// TwinCAT 3 PLC project Untitled1
// ProgramVersion: 3.1.4026.25
// libraries:
//   Tc2_Standard, * (Beckhoff Automation GmbH)
//   Tc2_System, * (Beckhoff Automation GmbH)
// project tree:
//   GVLs/ GVL.TcGVL
//   / PlcTask.TcTTO
//   POUs/ MAIN.TcPOU
// real-time tasks:
//   TASK PlcTask: cycle T#10ms, priority 20, ADS port 350
// motion (NC):
//   TASK NC-Task 1 SAF: cycle T#2ms, priority 4, ADS port 501
//   TASK NC-Task 1 SVB: cycle T#10ms, priority 8, ADS port 511
//   AXIS Axis 1 (id 1)
//     OtherSettings: AllowMotionCmdToSlave=true
//     encoder EncType=8
//       EncPara: MaxCount=#xffffffff
//     drive DrvType=9
//       DrvPara: MaxCount=#xffffffff, DriveControlDWord=#x00030000
//         Analog: VeloScale=6, TorqueSetpointScale=10, ScaleFactorActTorque=0.1
//         TimeComp: TaskDelayCycles=1
//     controller CtrType=1
//       CtrPara: PriorControlFactor=1
//         Observer: BandWidth=20
//   AXIS Axis 2 (id 2)
//     OtherSettings: AllowMotionCmdToSlave=true
//     encoder EncType=8
//       EncPara: MaxCount=#xffffffff
//     drive DrvType=9
//       DrvPara: MaxCount=#xffffffff, DriveControlDWord=#x00030000
//         Analog: VeloScale=6, TorqueSetpointScale=10, ScaleFactorActTorque=0.1
//         TimeComp: TaskDelayCycles=1
//     controller CtrType=1
//       CtrPara: PriorControlFactor=1
//         Observer: BandWidth=20
// I/O:
//   DEVICE Device 1 (EtherCAT), AmsNetId 192.168.0.5.2.1
//     Box 1 (CU1128) [CU1128 6x EtherCAT junction]
//       Box 10 (EP1018-0001) [EP1018-0001 8 Ch. Dig. Input 24V, 10µs, M8]
//       Box 11 (EP1018-0001) [EP1018-0001 8 Ch. Dig. Input 24V, 10µs, M8]
//       Box 12 (EP1018-0001) [EP1018-0001 8 Ch. Dig. Input 24V, 10µs, M8]
//       Box 13 (EP2028-0001) [EP2028-0001 8 Ch. Dig. Output 24V, 2A, M8]
//       Box 14 (EP2028-0001) [EP2028-0001 8 Ch. Dig. Output 24V, 2A, M8]
//       Term 7 (EK1100-0030) [EK1100-0030 EtherCAT Coupler (2A E-Bus, 4kV galv. iso.)]
//         Term 8 (EL1809) [EL1809 16Ch. Dig. Input 24V, 3ms]
//         Term 9 (EL2809) [EL2809 16Ch. Dig. Output 24V, 0.5A]
//       Term 4 (EK1100-0030) [EK1100-0030 EtherCAT Coupler (2A E-Bus, 4kV galv. iso.)]
//         Term 5 (EL1809) [EL1809 16Ch. Dig. Input 24V, 3ms]
//         Term 6 (EL2809) [EL2809 16Ch. Dig. Output 24V, 0.5A]
//         Drive 15 (AX5206-0000-0011) [AX5206-0000-0011 EtherCAT Drive (SoE, 2 Ch.)]
//       Box 2 (CU1128-B) [CU1128 6x EtherCAT junction - Dev A]
//       Box 3 (CU1128-C) [CU1128 6x EtherCAT junction - Dev B]
// variable links:
//   NC-Task 1 SAF/Axes/Axis 1 <-> Device 1 (EtherCAT)/Box 1 (CU1128)/Term 4 (EK1100-0030)/Drive 15 (AX5206-0000-0011)
//     Drive/Inputs/In/nDcOutputTime <-> InfoData/DcOutputShift
//     Drive/Inputs/In/nState1 <-> AT 1/Drive status word @bit 8
//     Drive/Inputs/In/nState2 <-> AT 1/Drive status word
//     Drive/Inputs/In/nState4 @bit 1 <-> WcState/InputToggle
//     Drive/Inputs/In/nState4 <-> WcState/WcState
//     Drive/Outputs/Out/nCtrl1 <-> MDT 1/Master control word @bit 8
//     Drive/Outputs/Out/nDataOut2 <-> MDT 1/Velocity command value
//     Enc/Inputs/In/nDataIn1 <-> AT 1/Position feedback 1 value
//     Enc/Inputs/In/nDcInputTime <-> InfoData/DcInputShift
//     Enc/Inputs/In/nState4 @bit 1 <-> WcState/InputToggle
//     Enc/Inputs/In/nState4 <-> WcState/WcState
//   NC-Task 1 SAF/Axes/Axis 2 <-> Device 1 (EtherCAT)/Box 1 (CU1128)/Term 4 (EK1100-0030)/Drive 15 (AX5206-0000-0011)
//     Drive/Inputs/In/nDcOutputTime <-> InfoData/DcOutputShift
//     Drive/Inputs/In/nState1 <-> AT 2/Drive status word @bit 8
//     Drive/Inputs/In/nState2 <-> AT 2/Drive status word
//     Drive/Inputs/In/nState4 @bit 1 <-> WcState/InputToggle
//     Drive/Inputs/In/nState4 <-> WcState/WcState
//     Drive/Outputs/Out/nCtrl1 <-> MDT 2/Master control word @bit 8
//     Drive/Outputs/Out/nDataOut2 <-> MDT 2/Velocity command value
//     Enc/Inputs/In/nDataIn1 <-> AT 2/Position feedback 1 value
//     Enc/Inputs/In/nDcInputTime <-> InfoData/DcInputShift
//     Enc/Inputs/In/nState4 @bit 1 <-> WcState/InputToggle
//     Enc/Inputs/In/nState4 <-> WcState/WcState
//   Untitled1/Untitled1 Instance <-> Device 1 (EtherCAT)/Box 1 (CU1128)/Box 10 (EP1018-0001)
//     PlcTask Inputs/GVL.bZylAuswerferAS <-> Channel 1/Input
//     PlcTask Inputs/GVL.bZylAuswerferGS <-> Channel 2/Input
//     PlcTask Inputs/GVL.bZylSpannerAS <-> Channel 3/Input
//     PlcTask Inputs/GVL.bZylSpannerGS <-> Channel 4/Input
//     PlcTask Inputs/GVL.bZylWeicheAS <-> Channel 5/Input
//     PlcTask Inputs/GVL.bZylWeicheGS <-> Channel 6/Input
//   Untitled1/Untitled1 Instance <-> Device 1 (EtherCAT)/Box 1 (CU1128)/Box 11 (EP1018-0001)
//     PlcTask Inputs/GVL.bZylAuslaufAS <-> Channel 3/Input
//     PlcTask Inputs/GVL.bZylAuslaufGS <-> Channel 4/Input
//     PlcTask Inputs/GVL.bZylEinlaufAS <-> Channel 1/Input
//     PlcTask Inputs/GVL.bZylEinlaufGS <-> Channel 2/Input
//   Untitled1/Untitled1 Instance <-> Device 1 (EtherCAT)/Box 1 (CU1128)/Box 12 (EP1018-0001)
//     PlcTask Inputs/GVL.bLS_Auslauf <-> Channel 5/Input
//     PlcTask Inputs/GVL.bLS_Einlauf <-> Channel 1/Input
//     PlcTask Inputs/GVL.bServoAuslaufAS <-> Channel 7/Input
//     PlcTask Inputs/GVL.bServoAuslaufGS <-> Channel 8/Input
//     PlcTask Inputs/GVL.bServoAuslaufRast <-> Channel 6/Input
//     PlcTask Inputs/GVL.bServoEinlaufAS <-> Channel 3/Input
//     PlcTask Inputs/GVL.bServoEinlaufGS <-> Channel 4/Input
//     PlcTask Inputs/GVL.bServoEinlaufRast <-> Channel 2/Input
//   Untitled1/Untitled1 Instance <-> Device 1 (EtherCAT)/Box 1 (CU1128)/Box 13 (EP2028-0001)
//     PlcTask Outputs/GVL.bVentilAuswerferAS <-> Channel 1/Output
//     PlcTask Outputs/GVL.bVentilAuswerferGS <-> Channel 2/Output
//     PlcTask Outputs/GVL.bVentilSpannerAS <-> Channel 3/Output
//     PlcTask Outputs/GVL.bVentilSpannerGS <-> Channel 4/Output
//     PlcTask Outputs/GVL.bVentilWeicheAS <-> Channel 5/Output
//     PlcTask Outputs/GVL.bVentilWeicheGS <-> Channel 6/Output
//   Untitled1/Untitled1 Instance <-> Device 1 (EtherCAT)/Box 1 (CU1128)/Box 14 (EP2028-0001)
//     PlcTask Outputs/GVL.bVentilAusblasenAS <-> Channel 5/Output
//     PlcTask Outputs/GVL.bVentilAusblasenGS <-> Channel 6/Output
//     PlcTask Outputs/GVL.bVentilAuslaufAS <-> Channel 3/Output
//     PlcTask Outputs/GVL.bVentilAuslaufGS <-> Channel 4/Output
//     PlcTask Outputs/GVL.bVentilAuswurfBypAS <-> Channel 7/Output
//     PlcTask Outputs/GVL.bVentilAuswurfBypGS <-> Channel 8/Output
//     PlcTask Outputs/GVL.bVentilEinlaufAS <-> Channel 1/Output
//     PlcTask Outputs/GVL.bVentilEinlaufGS <-> Channel 2/Output
//   Untitled1/Untitled1 Instance <-> Device 1 (EtherCAT)/Box 1 (CU1128)/Term 4 (EK1100-0030)/Term 5 (EL1809)
//     PlcTask Inputs/GVL.bDruckschalter <-> Channel 1/Input
//     PlcTask Inputs/GVL.bNotHalt <-> Channel 2/Input
//   Untitled1/Untitled1 Instance <-> Device 1 (EtherCAT)/Box 1 (CU1128)/Term 4 (EK1100-0030)/Term 6 (EL2809)
//     PlcTask Outputs/GVL.bEntlueften <-> Channel 1/Output
//     PlcTask Outputs/GVL.bLaserEnable <-> Channel 2/Output
//   Untitled1/Untitled1 Instance <-> Device 1 (EtherCAT)/Box 1 (CU1128)/Term 7 (EK1100-0030)/Term 8 (EL1809)
//     PlcTask Inputs/GVL.bCW_Adb_coded <-> Channel 2/Input
//     PlcTask Inputs/GVL.bCW_Eready <-> Channel 1/Input
//     PlcTask Inputs/GVL.bCW_MarkInProgress <-> Channel 3/Input
//   Untitled1/Untitled1 Instance <-> Device 1 (EtherCAT)/Box 1 (CU1128)/Term 7 (EK1100-0030)/Term 9 (EL2809)
//     PlcTask Outputs/GVL.bCW_ERR_RESET <-> Channel 2/Output
//     PlcTask Outputs/GVL.bCW_Ex_GO <-> Channel 1/Output
//     PlcTask Outputs/GVL.bCW_STAT_REQ <-> Channel 4/Output
//     PlcTask Outputs/GVL.bCW_STOP <-> Channel 3/Output

CONFIGURATION Untitled1
    RESOURCE PLC ON TwinCAT3
        TASK PlcTask(INTERVAL := T#10ms, PRIORITY := 20);
        PROGRAM MAIN WITH PlcTask : MAIN;
    END_RESOURCE
END_CONFIGURATION

// ---- GVLs/GVL.TcGVL
{attribute 'qualified_only'}
VAR_GLOBAL
    // ==========================================
    // MAIN CONTROL CABINET (Schaltschrank)
    // ==========================================
    
    // Inputs (EL1809 - +MP-6K10)
    bDruckschalter         AT %I* : BOOL; // E0.0 Wartungseinheit Druckschalter[cite: 15, 25]
    bNotHalt               AT %I* : BOOL; // E0.1 Not-Halt betätigt[cite: 15, 18]
    
    // Outputs (EL2809 - +MP-6K20)
    bEntlueften            AT %Q* : BOOL; // A0.0 Wartungseinheit Entlüften[cite: 15, 25]
    bLaserEnable           AT %Q* : BOOL; // A0.1 LaserEnable[cite: 15, 18]

    // ==========================================
    // CW CONTROLLER
    // ==========================================
    
    // Inputs (EL1809 - +LS-7K10)
    bCW_Eready             AT %I* : BOOL; // E50.0 CW Eready[cite: 17]
    bCW_Adb_coded          AT %I* : BOOL; // E50.1 CW Adb coded[cite: 17]
    bCW_MarkInProgress     AT %I* : BOOL; // E50.2 CW MarkInProgress[cite: 17]
    
    // Outputs (EL2809 - +LS-7K20)
    bCW_Ex_GO              AT %Q* : BOOL; // A50.0 CW Ex.GO[cite: 17]
    bCW_ERR_RESET          AT %Q* : BOOL; // A50.1 CW ERR_RESET[cite: 17]
    bCW_STOP               AT %Q* : BOOL; // A50.2 CW STOP[cite: 17]
    bCW_STAT_REQ           AT %Q* : BOOL; // A50.3 CW STAT_REQ[cite: 17]

    // ==========================================
    // FIELD BOX 1 (EP1018-0001 - +MS-9K1)
    // ==========================================
    
    bZylAuswerferAS        AT %I* : BOOL; // E1050.0 Zylinder Auswerfer AS (Port X1:4)[cite: 20, 30]
    bZylAuswerferGS        AT %I* : BOOL; // E1050.1 Zylinder Auswerfer GS (Port X2:4)[cite: 20, 30]
    bZylSpannerAS          AT %I* : BOOL; // E1050.2 Zylinder Spanner AS (Port X3:4)[cite: 20, 31]
    bZylSpannerGS          AT %I* : BOOL; // E1050.3 Zylinder Spanner GS (Port X4:4)[cite: 20, 31]
    bZylWeicheAS           AT %I* : BOOL; // E1050.4 Zylinder Weiche AS (Port X5:4)[cite: 20, 32]
    bZylWeicheGS           AT %I* : BOOL; // E1050.5 Zylinder Weiche GS (Port X6:4)[cite: 20, 32]

    // ==========================================
    // FIELD BOX 2 (EP1018-0001 - +MS-9K2)
    // ==========================================
    
    bZylEinlaufAS          AT %I* : BOOL; // E1051.0 Zylinder Einlauf AS (Port X1:4)[cite: 20, 27]
    bZylEinlaufGS          AT %I* : BOOL; // E1051.1 Zylinder Einlauf GS (Port X2:4)[cite: 20, 27]
    bZylAuslaufAS          AT %I* : BOOL; // E1051.2 Zylinder Auslauf AS (Port X3:4)[cite: 20, 29]
    bZylAuslaufGS          AT %I* : BOOL; // E1051.3 Zylinder Auslauf GS (Port X4:4)[cite: 20, 29]

    // ==========================================
    // FIELD BOX 3 (EP1018-0001 - +MS-9K3)
    // ==========================================
    
    bLS_Einlauf            AT %I* : BOOL; // E1052.0 Lichtschranke Einlauf (Port X1:4)[cite: 21, 26]
    bServoEinlaufRast      AT %I* : BOOL; // E1052.1 Servo Einlauf eingerastet (Port X2:4)[cite: 21, 26]
    bServoEinlaufAS        AT %I* : BOOL; // E1052.2 Servo Einlauf AS (Port X3:4)[cite: 21, 26]
    bServoEinlaufGS        AT %I* : BOOL; // E1052.3 Servo Einlauf GS (Port X4:4)[cite: 21, 26]
    bLS_Auslauf            AT %I* : BOOL; // E1052.4 Lichtschranke Auslauf (Port X5:4)[cite: 21, 28]
    bServoAuslaufRast      AT %I* : BOOL; // E1052.5 Servo Auslauf eingerastet (Port X6:4)[cite: 21, 28]
    bServoAuslaufAS        AT %I* : BOOL; // E1052.6 Servo Auslauf AS (Port X7:4)[cite: 21, 28]
    bServoAuslaufGS        AT %I* : BOOL; // E1052.7 Servo Auslauf GS (Port X8:4)[cite: 21, 28]

    // ==========================================
    // FIELD BOX 4 (EP2028-0001 - +MS-10K1)
    // ==========================================
    
    bVentilAuswerferAS     AT %Q* : BOOL; // A1050.0 Ventil Auswerfer AS (Port X1:4)[cite: 23, 30]
    bVentilAuswerferGS     AT %Q* : BOOL; // A1050.1 Ventil Auswerfer GS (Port X2:4)[cite: 23, 30]
    bVentilSpannerAS       AT %Q* : BOOL; // A1050.2 Ventil Spanner AS (Port X3:4)[cite: 23, 31]
    bVentilSpannerGS       AT %Q* : BOOL; // A1050.3 Ventil Spanner GS (Port X4:4)[cite: 23, 31]
    bVentilWeicheAS        AT %Q* : BOOL; // A1050.4 Ventil Weiche AS (Port X5:4)[cite: 23, 32]
    bVentilWeicheGS        AT %Q* : BOOL; // A1050.5 Ventil Weiche GS (Port X6:4)[cite: 23, 32]

    // ==========================================
    // FIELD BOX 5 (EP2028-0001 - +MS-10K2)
    // ==========================================
    
    bVentilEinlaufAS       AT %Q* : BOOL; // A1051.0 Ventil Einlauf AS (Port X1:4)[cite: 23, 27]
    bVentilEinlaufGS       AT %Q* : BOOL; // A1051.1 Ventil Einlauf GS (Port X2:4)[cite: 23, 27]
    bVentilAuslaufAS       AT %Q* : BOOL; // A1051.2 Ventil Auslauf AS (Port X3:4)[cite: 23, 29]
    bVentilAuslaufGS       AT %Q* : BOOL; // A1051.3 Ventil Auslauf GS (Port X4:4)[cite: 23, 29]
    bVentilAusblasenAS     AT %Q* : BOOL; // A1051.4 Ventil Ausblasen AS (Port X5:4)[cite: 23, 33]
    bVentilAusblasenGS     AT %Q* : BOOL; // A1051.5 Ventil Ausblasen GS (Port X6:4)[cite: 23, 33]
    bVentilAuswurfBypAS    AT %Q* : BOOL; // A1051.6 Ventil Auswurf Bypass AS (Port X7:4)[cite: 23, 34]
    bVentilAuswurfBypGS    AT %Q* : BOOL; // A1051.7 Ventil Auswurf Bypass GS (Port X8:4)[cite: 23, 34]
END_VAR

// ---- POUs/MAIN.TcPOU
PROGRAM MAIN
VAR
END_VAR

END_PROGRAM
